// TIA Portal V20 export
TYPE "WT3_Verbund_Status_UDT"
   STRUCT
      iHandshake : Int;
      Alarm : Struct
         bE0000_KonfigAlarm : Bool;
         bE0001_Reserviert : Bool;
         bE0002_InvUngueltig : Bool;
         bE0003_Reserviert : Bool;
         bE0004_Reserviert : Bool;
         bE0005_Reserviert : Bool;
         bE0006_Reserviert : Bool;
         bE0007_KonfigAlarmKdKonst : Bool;
         bE0008_KonfigAlarmVrKonst : Bool;
         bE0009_Reserviert : Bool;
         bE0010_Reserviert : Bool;
         bE0011_Reserviert : Bool;
         bE0012_Reserviert : Bool;
         bE0013_HdVerbundLäuftNicht : Bool;
         bE0014_HdVerbundLäuftNicht : Bool;
         b037_Reserve : Bool;
         by04_Reserve : Byte;
         by05_Reserve : Byte;
         by06_Reserve : Byte;
         by07_Reserve : Byte;
         by08_Reserve : Byte;
         by09_Reserve : Byte;
         by10_Reserve : Byte;
         by11_Reserve : Byte;
         by12_Reserve : Byte;
         by13_Reserve : Byte;
         by14_Reserve : Byte;
         by15_Reserve : Byte;
         by16_Reserve : Byte;
         by17_Reserve : Byte;
         by18_Reserve : Byte;
         by19_Reserve : Byte;
         by20_Reserve : Byte;
         by21_Reserve : Byte;
         by22_Reserve : Byte;
         by23_Reserve : Byte;
         by24_Reserve : Byte;
         by25_Reserve : Byte;
         by26_Reserve : Byte;
         bE0200_AlarmKabelbruch : Bool;
         b271_Reserve : Bool;
         b272_Reserve : Bool;
         b273_Reserve : Bool;
         b274_Reserve : Bool;
         b275_Reserve : Bool;
         b276_Reserve : Bool;
         b277_Reserve : Bool;
         by28_Reserve : Byte;
         by29_Reserve : Byte;
         by30_Reserve : Byte;
         by31_Reserve : Byte;
         by32_Reserve : Byte;
         by33_Reserve : Byte;
      END_STRUCT;
      Warnung : Struct
         bA1000_Reserviert : Bool;
         bA1001_SlaveAusg : Bool;
         bA1002_Reserviert : Bool;
         bA1003_HauptMasterAusg : Bool;
         bA1004_ZuwenigVDLeistungVerf : Bool;
         bA1005_HDVerbundAusg : Bool;
         bA1006_NDVerbundAusg : Bool;
         bA1007_Reserviert : Bool;
         bA1008_Reserviert : Bool;
         bA1009_MVbMasterAktiv : Bool;
         bA1010_ObjektIDMehrfVorhanden : Bool;
         b1011_KonfigWarnungAnfVd : Bool;
         b1012_KonfigWarnungFreigabeVd : Bool;
         b355_Reserve : Bool;
         b356_Reserve : Bool;
         b357_Reserve : Bool;
         by36_Reserve : Byte;
         by37_Reserve : Byte;
         by38_Reserve : Byte;
         by39_Reserve : Byte;
         by40_Reserve : Byte;
         by41_Reserve : Byte;
         by42_Reserve : Byte;
         by43_Reserve : Byte;
         by44_Reserve : Byte;
         by45_Reserve : Byte;
         by46_Reserve : Byte;
         by47_Reserve : Byte;
         by48_Reserve : Byte;
         by49_Reserve : Byte;
         by50_Reserve : Byte;
         by51_Reserve : Byte;
         by52_Reserve : Byte;
         by53_Reserve : Byte;
         by54_Reserve : Byte;
         by55_Reserve : Byte;
         by56_Reserve : Byte;
         by57_Reserve : Byte;
         by58_Reserve : Byte;
         bA1200_WarnungKabelbruch : Bool;
         b591_Reserve : Bool;
         b592_Reserve : Bool;
         b593_Reserve : Bool;
         b594_Reserve : Bool;
         b595_Reserve : Bool;
         b596_Reserve : Bool;
         b597_Reserve : Bool;
         by60_Reserve : Byte;
         by61_Reserve : Byte;
         by62_Reserve : Byte;
         by63_Reserve : Byte;
         by64_Reserve : Byte;
         by65_Reserve : Byte;
      END_STRUCT;
      Zustand : Struct
         bAlarmzustandAktiv : Bool;
         bWarnzustandAktiv : Bool;
         bSystemMeldungAktiv : Bool;
         bSeviceMeldungAktiv : Bool;
         bStopManuell : Bool;
         bStopAuto : Bool;
         bStopExtern : Bool;
         bBetriebAuto : Bool;
         bBetriebManuell : Bool;
         bAnlaufAuto : Bool;
         bAnlaufManuell : Bool;
         bManuellStoppen : Bool;
         b674_Reserve : Bool;
         b675_Reserve : Bool;
         b676_Reserve : Bool;
         b677_Reserve : Bool;
         by68_Reserve : Byte;
         by69_Reserve : Byte;
         bInventarAufnahme : Bool;
         bStartbefehlManuell : Bool;
         bStandbyMasterInit : Bool;
         bStandbyMasterPassiv : Bool;
         bStandbyMasterAktiv : Bool;
         bInitialisierung : Bool;
         bFreigabeWeitVdNötig : Bool;
         bAnforderungVdAktiv : Bool;
         bZuschSperreTodband : Bool;
         bBeschrLaufendeVd : Bool;
         bZuschSperreSinkenderBed : Bool;
         bLastsperreAktiv : Bool;
         bMasterGesperrt : Bool;
         bSollwertAnhebung : Bool;
         bSollwertAbsenkung : Bool;
         bPSaugTiefSperre : Bool;
         bAnfHDVerbund : Bool;
         bBoosterFreigabeFehlt : Bool;
         bAnforderungBooster : Bool;
         bHDVerbundFreigabeFehlt : Bool;
         bHDVerbundFreigabeMan : Bool;
         bBoosterFreigabeMan : Bool;
         bLeistBeschrAktiv : Bool;
         bZuschSperreLeistBesch : Bool;
         bZuschaltverzögerung : Bool;
         bPDruckLimitAktiv : Bool;
         bPSaugLimitaktiv : Bool;
         bPDruckGradLimitAktiv : Bool;
         bPSaugGradLimitAktiv : Bool;
         bVerbundRampeAktiv : Bool;
         bVetoReglerAktiv : Bool;
         b737_Reserve : Bool;
         by74_Reserve : Byte;
         by75_Reserve : Byte;
         by76_Reserve : Byte;
         by77_Reserve : Byte;
         by78_Reserve : Byte;
         by79_Reserve : Byte;
         by80_Reserve : Byte;
         by81_Reserve : Byte;
      END_STRUCT;
      "Allgemeine Meldungen" : Struct
         b4000_AllgemeineMeldung_1 : Bool;
         b4001_AllgemeineMeldung_2 : Bool;
         b4002_AllgemeineMeldung_3 : Bool;
         b4003_AllgemeineMeldung_4 : Bool;
         b4004_AllgemeineMeldung_5 : Bool;
         b4005_AllgemeineMeldung_6 : Bool;
         b4006_AllgemeineMeldung_7 : Bool;
         b4007_AllgemeineMeldung_8 : Bool;
         by83_Reserve : Byte;
         by84_Reserve : Byte;
         by85_Reserve : Byte;
      END_STRUCT;
      DigIn : Struct
         bStartbefehlVerbund : Bool;
         bSollwertB : Bool;
         bVerbundleistExtPlus : Bool;
         bVerbundleistExtMinus : Bool;
         bElLeistungZuHoch : Bool;
         bSollwertBHeizen : Bool;
         bUmschaltungWirksinn : Bool;
         b867_Reserve : Bool;
         by87_Reserve : Byte;
         by88_Reserve : Byte;
         by89_Reserve : Byte;
         by90_Reserve : Byte;
         by91_Reserve : Byte;
         by92_Reserve : Byte;
         by93_Reserve : Byte;
      END_STRUCT;
      DigOut : Struct
         bVerbundBereit : Bool;
         b941_Reserve : Bool;
         bFreigabeBoosterVerbund : Bool;
         bWarnungVerfuegbareLeistung : Bool;
         b944_Reserve : Bool;
         b945_Reserve : Bool;
         b946_Reserve : Bool;
         b947_Reserve : Bool;
         by95_Reserve : Byte;
         by96_Reserve : Byte;
         by97_Reserve : Byte;
         by98_Reserve : Byte;
         by99_Reserve : Byte;
         by100_Reserve : Byte;
         by101_Reserve : Byte;
      END_STRUCT;
      iAnzVd : Int;
      chRemoteSensEinheit : Char;
      chLeistRegEinheit : Char;
      rLeistRegIst : Real;
      rLeistRegSoll : Real;
      rVerbLeistSoll : Real;
      rVerbLeistSollVol : Real;
      rVerbLeistIst : Real;
      rVerbLeistIstVol : Real;
      rVeV : Real;
      rVevVol : Real;
      rVeD : Real;
      rVedVol : Real;
      rFVolMaxVerbund : Real;
      iNaechsterVdein : Int;
      iNaechsterVdaus : Int;
      rRemoteSensIst : Real;
      rVrTempEin : Real;
      rVrTempAus : Real;
      rKdrTempEin : Real;
      rKdrTempAus : Real;
      diStatusSollwertRampe : DInt;
      rRegelabweichungProz : Real;
      rRegelabweichung : Real;
      rReglerSollwertHeizenProz : Real;
      rReglerSollwertHeizen : Real;
      diStatussollwertrampeHeizen : DInt;
      rReglerIstwertheizenProz : Real;
      rReglerIstwertHeizen : Real;
      rRegelabweichungHeizenProz : Real;
      rRegelabweichungHeizen : Real;
      rVetoLimitProz : Real;
      rVetoLimit : Real;
      diNächsterVdEin : DInt;
      rVerbundleistungVdEin : Real;
      diNächsterVdAus : DInt;
      rVerbundleistungVdAus : Real;
      rLeistungslimitExternFeldbus : Real;
      rLeistungslimitExternAnalog : Real;
      rLeistungsbeschränkungMax : Real;
      rPDruckseite : Real;
      rPDuckseitetemp : Real;
      rPSaugseite : Real;
      rPSaugseiteTemp : Real;
      rRemoteIstwertHeizen : Real;
      rAuxAnalog1 : Real;
      rAuxAnalog2 : Real;
      rAnalogeLeistungsbeschränkung : Real;
      byReserve : Array[282..629] of Byte;
   END_STRUCT;
END_TYPE
